Staubli VAL3: if_check.pgx

public program if_check(num x_nType, num x_nIndex, num x_nValue, bool& x_bResult, bool& x_bDisable)
  local bool l_bErr
  local bool l_bValue
  local bool l_bRecValue
  local num l_nRecValue
begin
   x_bDisable=false
    switch x_nType
      case 1
        //din
        call io:getDigIO(io:dInput[x_nIndex],l_bRecValue,l_bErr)
        l_bValue=(x_nValue!=0)
        x_bResult=(l_bRecValue==l_bValue)
      break
      case 2
        //dout
        call io:getDigIO(io:dOutput[x_nIndex],l_bRecValue,l_bErr)
        l_bValue=(x_nValue!=0)
        x_bResult=(l_bRecValue==l_bValue)
      break
      case 3
        //ain
        call io:getAnaIO(io:aInput[x_nIndex],l_nRecValue,l_bErr)
        x_bResult=(l_nRecValue==x_nValue)
      break
      case 4
        //aout
        call io:getAnaIO(io:aInput[x_nIndex],l_nRecValue,l_bErr)
        x_bResult=(l_nRecValue==x_nValue)
      break
    default
      x_bDisable=true
    break
    endSwitch

end
